Staubli VAL3: computeZone.pgx

public program computeZone(num x_nIndex, bool& x_bResult)
  local tool l_tTool
  local frame l_fFrame
  local trsf l_trFirst
  local trsf l_trSecond
  local num l_nMax_x
  local num l_nMax_y
  local num l_nMax_z
  local num l_nMin_x
  local num l_nMin_y
  local num l_nMin_z
  local pointRx l_pPoint
  local bool l_bReuslt1
  local bool l_bReuslt2
  local bool l_bReuslt3
begin
  link(l_tTool,flange)
  link(l_fFrame,world)
  l_fFrame.trsf=safeTemp:zZoneItem[x_nIndex].fBase.trsf
  call savedata:getTool(nToolIndex,l_tTool)
  l_pPoint=here(l_tTool,l_fFrame)
  l_trFirst=safeTemp:zZoneItem[x_nIndex].pFirst.trsf
  l_trSecond=safeTemp:zZoneItem[x_nIndex].pSecond.trsf

  l_nMax_x=max(l_trFirst.x,l_trSecond.x)
  l_nMax_y=max(l_trFirst.y,l_trSecond.y)
  l_nMax_z=max(l_trFirst.z,l_trSecond.z)
  l_nMin_x=min(l_trFirst.x,l_trSecond.x)
  l_nMin_y=min(l_trFirst.y,l_trSecond.y)
  l_nMin_z=min(l_trFirst.z,l_trSecond.z)

  if l_nMin_x<l_pPoint.trsf.x and l_pPoint.trsf.x<l_nMax_x
    l_bReuslt1=true
  else
    l_bReuslt1=false
  endIf

  if l_nMin_y<l_pPoint.trsf.y and l_pPoint.trsf.y<l_nMax_y
    l_bReuslt2=true
  else
    l_bReuslt2=false
  endIf

  if l_nMin_z<l_pPoint.trsf.z and l_pPoint.trsf.z<l_nMax_z
    l_bReuslt3=true
  else
    l_bReuslt3=false
  endIf

  if l_bReuslt1 and l_bReuslt2 and l_bReuslt3
    x_bResult=true
  else
    x_bResult=false
  endIf
end
